// TIA Portal V21 export
FUNCTION_BLOCK "TiaMcpComponentGate"   // FB2, SCL
{ S7_Optimized_Access := 'TRUE' }
// stored: AutoNumber true, IsIECCheckEnabled false, IsRetainMemResEnabled false, MemoryReserve 100, SetENOAutomatically false, UDAEnableTagReadback false
   VAR_INPUT
      Enable : Bool;
   END_VAR
   VAR_OUTPUT
      Active : Bool;
   END_VAR
   VAR
      State { S7_SetPoint := 'True'} : "TiaMcpComponentState";
   END_VAR
BEGIN

       #State.Active := #Enable;
       #Active := #State.Active;
END_FUNCTION_BLOCK
